// TIA Portal V20 export
ORGANIZATION_BLOCK "Main"   // OB1, LAD, ProgramCycle
TITLE = "Main Program Sweep (Cycle)"
{ S7_Optimized_Access := 'TRUE' }
// stored: SetENOAutomatically false
   VAR_INPUT
      Initial_Call : Bool;   // Initial call of this OB
      Remanence : Bool;   // =True, if remanent data are available
   END_VAR
BEGIN

REGION Network 1
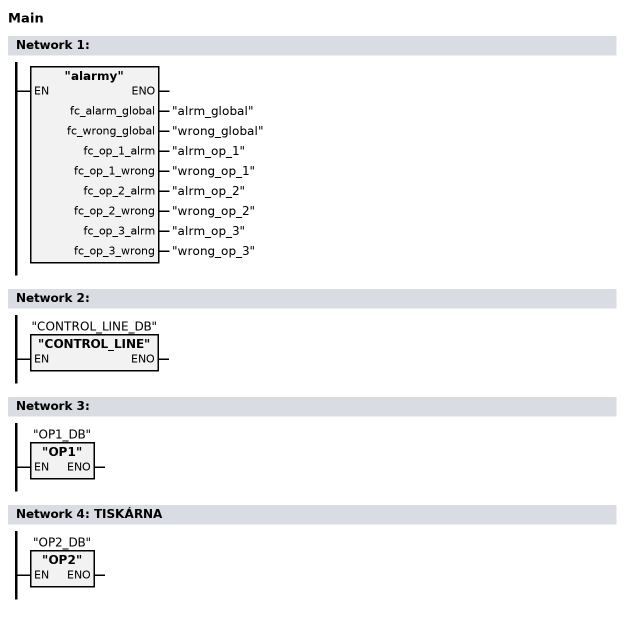
   RUNG wire#powerrail
      "alarmy"(fc_alarm_global => "alrm_global", fc_wrong_global => "wrong_global", fc_op_1_alrm => "alrm_op_1", fc_op_1_wrong => "wrong_op_1", fc_op_2_alrm => "alrm_op_2", fc_op_2_wrong => "wrong_op_2", fc_op_3_alrm => "alrm_op_3", fc_op_3_wrong => "wrong_op_3")
   END_RUNG
   // the same network as SCL:
   "alarmy"(fc_alarm_global => "alrm_global",
            fc_wrong_global => "wrong_global",
            fc_op_1_alrm => "alrm_op_1",
            fc_op_1_wrong => "wrong_op_1",
            fc_op_2_alrm => "alrm_op_2",
            fc_op_2_wrong => "wrong_op_2",
            fc_op_3_alrm => "alrm_op_3",
            fc_op_3_wrong => "wrong_op_3");
END_REGION

REGION Network 2
   RUNG wire#powerrail
      "CONTROL_LINE_DB"()
   END_RUNG
   // the same network as SCL:
   "CONTROL_LINE_DB"();   // "CONTROL_LINE"
END_REGION

REGION Network 3
   RUNG wire#powerrail
      "OP1_DB"()
   END_RUNG
   // the same network as SCL:
   "OP1_DB"();   // "OP1"
END_REGION

REGION Network 4: TISKÁRNA
   RUNG wire#powerrail
      "OP2_DB"()
   END_RUNG
   // the same network as SCL:
   "OP2_DB"();   // "OP2"
END_REGION
END_ORGANIZATION_BLOCK
